// TIA Portal V21 export
// export: Created 2026-11-08T21:35:20.4632136Z, ExportSetting WithDefaults, DisplayName Totally Integrated Automation Portal, DisplayVersion V21 Update 3, DisplayName STEP 7 Professional, DisplayVersion V21 Update 3, DisplayName STEP 7 Safety, DisplayVersion V21, DisplayName Tech WebApplication, DisplayVersion V21, DisplayName WinCC Basic/Comfort/Advanced, DisplayVersion V21 Update 3, DisplayName WinCC Unified, DisplayVersion V21 Update 3
FUNCTION_BLOCK "FB_StlC_012"   // FB89, STL
TITLE = STL call CompType
{ S7_Optimized_Access := 'TRUE' }
VERSION : 0.1
// stored: AutoNumber true, IsRetainMemResEnabled false, MemoryReserve 100, UDAEnableTagReadback false
   VAR_OUTPUT
      "b" : Bool;
   END_VAR
   VAR
      a1 : Array[0..3] of Int;
      a2 : Array[0..3] of Int;
   END_VAR
BEGIN

NETWORK
TITLE = 012 CompType
      CALL  CompType
      ( IN1 := #a1,
        IN2 := #a2,
        OUT := #"b"
      );
END_FUNCTION_BLOCK
